(* IEC 61131-3 sources: kns-pump-station/tests/POUs/Field/FB_VfdAdapter_Cond_Test, 9 files *)

(* ---- FB_VfdAdapter_Cond_Test.decl.st ---- *)
// Назначение: набор coUnit для FB_VfdAdapter_Cond — условная карта ПЧ: биты слова состояния, масштаб
//             частоты (5000 = 100 %), потеря связи (статусы FALSE, скорость удерживается), бит сброса в
//             слове управления, задание частоты с ограничением, округлением и защитой от NaN.
// Автор:      kr0nsch
// Версия:     0.1.0
// Документ:   docs/DESIGN.md, разделы 8.2, 14.1
FUNCTION_BLOCK FB_VfdAdapter_Cond_Test EXTENDS coUnit.FB_TestSuite
VAR CONSTANT
    R_EPS_PCT : REAL := 1.0E-4;     // допуск сравнения скорости, %
END_VAR

(* ---- DecodeBits.method.decl.st ---- *)
// Биты STW.0…STW.4 при связи: готов, в работе, авария, предупреждение, управление от клемм — каждый в свой
// выход; два разных слова проверяют, что биты не перепутаны
METHOD PRIVATE DecodeBits
VAR
    fbDut : FB_VfdAdapter_Cond;     // проверяемый адаптер
END_VAR

(* ---- DecodeScale5000Is100Pct.method.decl.st ---- *)
// Фактическая частота 0,01 Гц: 5000 → 100 %, 2500 → 50 %, 1 → 0,02 %
METHOD PRIVATE DecodeScale5000Is100Pct
VAR
    fbDut : FB_VfdAdapter_Cond;     // проверяемый адаптер
END_VAR

(* ---- DefaultsAllFalse.method.decl.st ---- *)
// Новый адаптер: связи нет, статусы FALSE, скорость, слово управления и задание — 0
METHOD PRIVATE DefaultsAllFalse
VAR
    fbDut : FB_VfdAdapter_Cond;     // проверяемый адаптер
END_VAR

(* ---- EncodeNanIsZero.method.decl.st ---- *)
// Неконечное задание (NaN, +Inf) — 0; бит сброса от задания не зависит
METHOD PRIVATE EncodeNanIsZero
VAR
    fbDut : FB_VfdAdapter_Cond;     // проверяемый адаптер
    uBits : PL.U_RealBits;          // сборка NaN и бесконечности из битов
END_VAR

(* ---- EncodeResetBitWhileQReset.method.decl.st ---- *)
// Слово управления: бит сброса аварии (CTW.2), пока есть импульс xQReset; бит пуска не используется
METHOD PRIVATE EncodeResetBitWhileQReset
VAR
    fbDut : FB_VfdAdapter_Cond;     // проверяемый адаптер
END_VAR

(* ---- EncodeRoundsToNearest.method.decl.st ---- *)
// Задание частоты округляется до ближайшего отсчёта 0,01 Гц, а не отбрасывается дробная часть:
// 12,358 % → 617,9 → 618; 12,342 % → 617,1 → 617; 99,995 % → 4999,75 → 5000
METHOD PRIVATE EncodeRoundsToNearest
VAR
    fbDut : FB_VfdAdapter_Cond;     // проверяемый адаптер
END_VAR

(* ---- EncodeScaleAndClamp.method.decl.st ---- *)
// Задание частоты: 50 % → 2500, 12,345 % → 617 (округление), выше 100 % → 5000, ниже 0 → 0, 100 % → 5000
METHOD PRIVATE EncodeScaleAndClamp
VAR
    fbDut : FB_VfdAdapter_Cond;     // проверяемый адаптер
END_VAR

(* ---- NoCommForcesStatusFalseHoldsSpeed.method.decl.st ---- *)
// Нет связи: регистры недостоверны — статусы FALSE (в том числе авария), скорость — последняя принятая (75 %);
// связь вернулась — снова по регистрам
METHOD PRIVATE NoCommForcesStatusFalseHoldsSpeed
VAR
    fbDut : FB_VfdAdapter_Cond;     // проверяемый адаптер
    wAll  : WORD;                   // все биты условной карты
END_VAR
